(* IEC 61131-3 sources: s7-to-codesys/src/POUs/S7Compat/F_NormX, 2 files *)

(* ---- F_NormX.decl.st ---- *)
// Назначение: аналог инструкции S7 NORM_X (S7-1200/1500) для кода, сконвертированного s7conv:
//             нормирование OUT = (VALUE - MIN) / (MAX - MIN). Значение вне MIN…MAX не
//             ограничивается: результат линейно продолжается ниже 0.0 и выше 1.0 (в S7 при этом
//             ENO = TRUE). При MIN > MAX — та же формула без перестановки границ; при MIN = MAX
//             результат 0.0 (деления на ноль нет). В S7 для MIN >= MAX ENO = FALSE, а значение
//             OUT не документировано — сверить с источником. ENO не воспроизводится.
// Автор:      kr0nsch
// Версия:     0.1.0
// Документ:   docs/MAPPING.md, раздел «NORM_X и SCALE_X»
FUNCTION F_NormX : REAL
VAR_INPUT
    rMin : REAL;        // нижняя граница диапазона значения (MIN в S7)
    rValue : REAL;      // нормируемое значение (VALUE в S7)
    rMax : REAL;        // верхняя граница диапазона значения (MAX в S7)
END_VAR
VAR
    rSpan : REAL;       // ширина диапазона MAX - MIN
END_VAR

(* ---- F_NormX.impl.st ---- *)
// Линейное нормирование без ограничения: вне MIN…MAX результат < 0.0 или > 1.0.
// Сравнение «больше или меньше» вместо «не равно»: проверка ширины диапазона без
// сравнения REAL на равенство.
IF rMax > rMin OR rMax < rMin THEN
    rSpan := rMax - rMin;
    F_NormX := (rValue - rMin) / rSpan;
ELSE
    // Вырожденный диапазон (в S7 — ENO = FALSE): делить на ноль нельзя, результат 0.0
    F_NormX := 0.0;
END_IF
